FUNCTION_BLOCK Basic1_1 (* Basic Function Block Type *)
  (* Standard: 61499-2 *)
  (* Version 0.0, 1/4/2020, prana, nxtControl GmbH, Template *)
  PACKAGE Main;
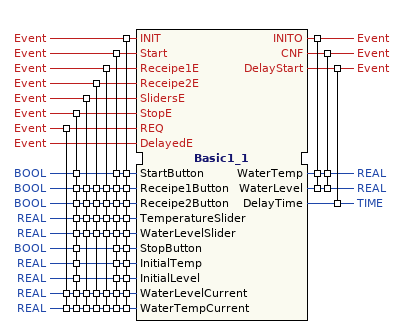
  EVENT_INPUT
    INIT WITH StartButton, Receipe1Button, Receipe2Button, TemperatureSlider, WaterLevelSlider, StopButton, InitialTemp, InitialLevel, WaterLevelCurrent, WaterTempCurrent;
    Start WITH StartButton, Receipe1Button, Receipe2Button, TemperatureSlider, WaterLevelSlider, StopButton, InitialTemp, InitialLevel, WaterLevelCurrent, WaterTempCurrent;
    Receipe1E WITH Receipe1Button, Receipe2Button, TemperatureSlider, WaterLevelSlider, WaterLevelCurrent, WaterTempCurrent; (* Initialization Request *)
    Receipe2E WITH Receipe1Button, Receipe2Button, TemperatureSlider, WaterLevelSlider, WaterLevelCurrent, WaterTempCurrent; (* Normal Execution Request *)
    SlidersE WITH Receipe1Button, Receipe2Button, TemperatureSlider, WaterLevelSlider, WaterLevelCurrent, WaterTempCurrent;
    StopE WITH StartButton, Receipe1Button, Receipe2Button, TemperatureSlider, WaterLevelSlider, StopButton, InitialTemp, InitialLevel, WaterLevelCurrent, WaterTempCurrent;
    REQ WITH WaterLevelCurrent, WaterTempCurrent;
    DelayedE;
  END_EVENT
  EVENT_OUTPUT
    INITO WITH WaterLevel, WaterTemp; (* Initialization Confirm *)
    CNF WITH WaterLevel, WaterTemp; (* Execution Confirmation *)
    DelayStart WITH DelayTime;
  END_EVENT
  VAR_INPUT
    StartButton : BOOL;
    Receipe1Button : BOOL; (* Input event qualifier *)
    Receipe2Button : BOOL;
    TemperatureSlider : REAL;
    WaterLevelSlider : REAL;
    StopButton : BOOL;
    InitialTemp : REAL;
    InitialLevel : REAL;
    WaterLevelCurrent : REAL;
    WaterTempCurrent : REAL;
  END_VAR
  VAR_OUTPUT
    WaterTemp : REAL;
    WaterLevel : REAL; (* Output event qualifier *)
    DelayTime : TIME;
  END_VAR
  VAR
    X1 : REAL := 160.50;
    Y1 : REAL := 50.00;
    X2 : REAL := 250.50;
    Y2 : REAL := 68.96;
    X3 : REAL := 351.50;
    Y3 : REAL := 64.32;
    X4 : REAL := 180.00;
    Y4 : REAL := 42.60;
    T1 : TIME := T#3s;
    T2 : TIME := T#2s;
  END_VAR
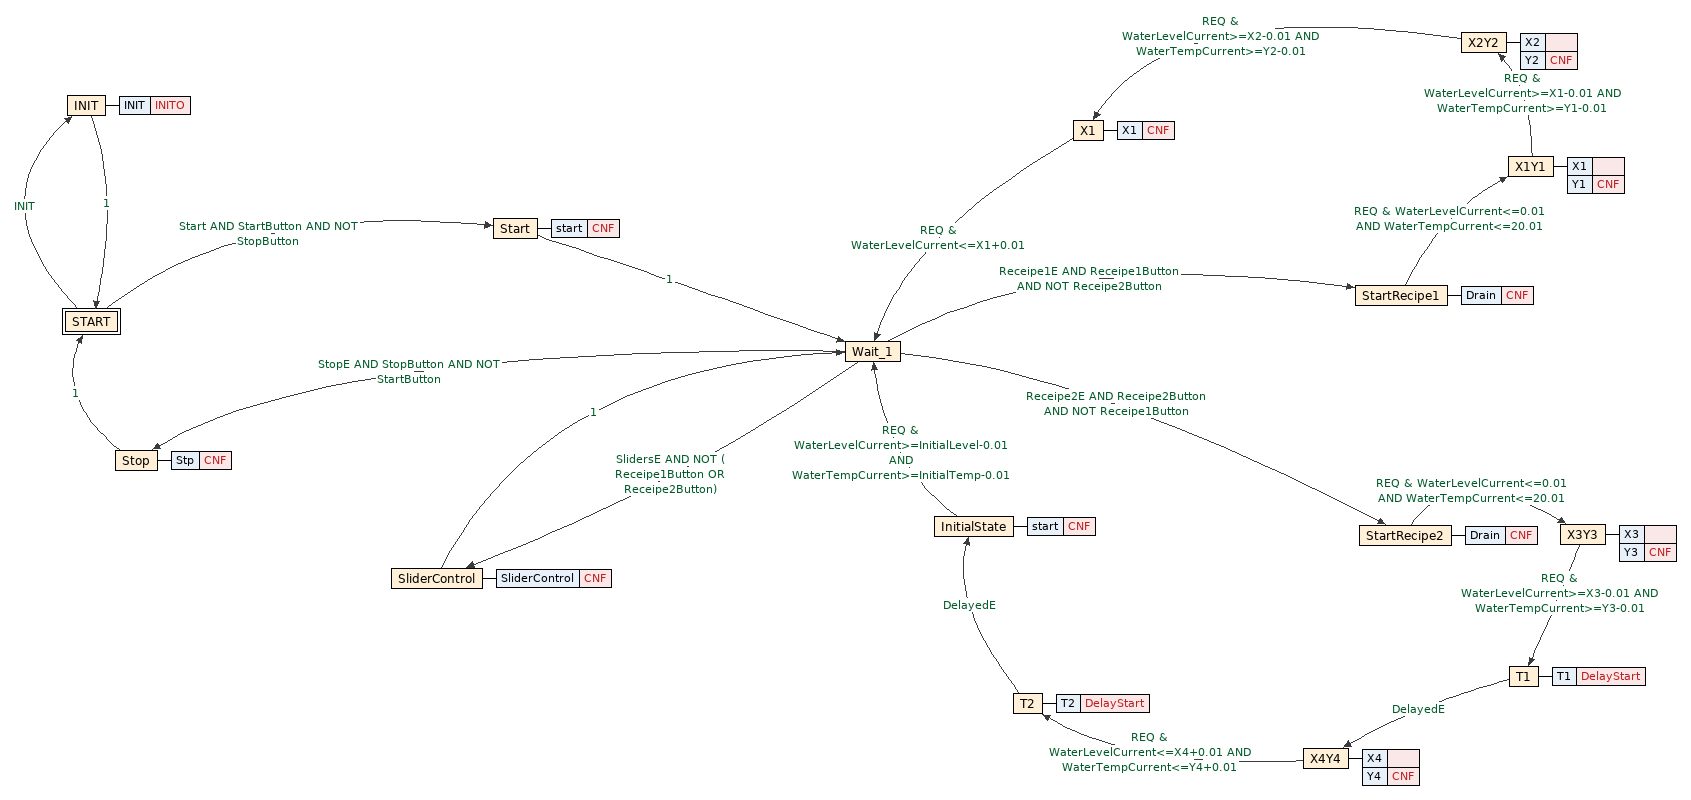
  EC_STATES
    START; (* Initial State *)
    SliderControl : SliderControl -> CNF;
    Start : start -> CNF;
    Wait_1;
    Stop : Stp -> CNF;
    INIT : INIT -> INITO;
    StartRecipe1 : Drain -> CNF;
    StartRecipe2 : Drain -> CNF;
    X1Y1 : X1, Y1 -> CNF;
    X2Y2 : X2, Y2 -> CNF;
    X1 : X1 -> CNF;
    X3Y3 : X3, Y3 -> CNF;
    T1 : T1 -> DelayStart;
    X4Y4 : X4, Y4 -> CNF;
    T2 : T2 -> DelayStart;
    InitialState : start -> CNF;
  END_STATES
  EC_TRANSITIONS
    Wait_1 TO SliderControl := SlidersE AND NOT ( Receipe1Button OR Receipe2Button);
    SliderControl TO Wait_1 := 1;
    START TO Start := Start AND StartButton AND NOT StopButton;
    Wait_1 TO Stop := StopE AND StopButton AND NOT StartButton;
    Stop TO START := 1;
    START TO INIT := INIT;
    INIT TO START := 1;
    StartRecipe1 TO X1Y1 := REQ & WaterLevelCurrent<=0.01 AND WaterTempCurrent<=20.01;
    X1Y1 TO X2Y2 := REQ & WaterLevelCurrent>=X1-0.01 AND WaterTempCurrent>=Y1-0.01;
    X3Y3 TO T1 := REQ & WaterLevelCurrent>=X3-0.01 AND WaterTempCurrent>=Y3-0.01;
    T1 TO X4Y4 := DelayedE;
    T2 TO InitialState := DelayedE;
    InitialState TO Wait_1 := REQ & WaterLevelCurrent>=InitialLevel-0.01 AND WaterTempCurrent>=InitialTemp-0.01;
    X2Y2 TO X1 := REQ & WaterLevelCurrent>=X2-0.01 AND WaterTempCurrent>=Y2-0.01;
    X1 TO Wait_1 := REQ & WaterLevelCurrent<=X1+0.01;
    Start TO Wait_1 := 1;
    Wait_1 TO StartRecipe1 := Receipe1E AND Receipe1Button AND NOT Receipe2Button;
    Wait_1 TO StartRecipe2 := Receipe2E AND Receipe2Button AND NOT Receipe1Button;
    StartRecipe2 TO X3Y3 := REQ & WaterLevelCurrent<=0.01 AND WaterTempCurrent<=20.01;
    X4Y4 TO T2 := REQ & WaterLevelCurrent<=X4+0.01 AND WaterTempCurrent<=Y4+0.01;
  END_TRANSITIONS
  ALGORITHM INIT IN ST: (* Initialization algorithm *)
;
  END_ALGORITHM
  ALGORITHM SliderControl IN ST:
WaterLevel := WaterLevelSlider;
WaterTemp := TemperatureSlider;
  END_ALGORITHM
  ALGORITHM start IN ST:
WaterLevel := InitialLevel;
WaterTemp := InitialTemp;
  END_ALGORITHM
  ALGORITHM Stp IN ST:
WaterLevel := 0;
WaterTemp := 0;
  END_ALGORITHM
  ALGORITHM Drain IN ST:
WaterLevel:=0;
WaterTemp:=0;
  END_ALGORITHM
  ALGORITHM X1 IN ST:
WaterLevel:=X1;
  END_ALGORITHM
  ALGORITHM Y1 IN ST:
WaterTemp:=Y1;
  END_ALGORITHM
  ALGORITHM X2 IN ST:
WaterLevel:=X2;
  END_ALGORITHM
  ALGORITHM Y2 IN ST:
WaterTemp:=Y2;
  END_ALGORITHM
  ALGORITHM X3 IN ST:
WaterLevel:=X3;
  END_ALGORITHM
  ALGORITHM X4 IN ST:
WaterLevel:=X4;
  END_ALGORITHM
  ALGORITHM Y3 IN ST:
WaterTemp:=Y3;
  END_ALGORITHM
  ALGORITHM Y4 IN ST:
WaterTemp:=Y4;
  END_ALGORITHM
  ALGORITHM T1 IN ST:
DelayTime:=T1;
  END_ALGORITHM
  ALGORITHM T2 IN ST:
DelayTime:=T2;
  END_ALGORITHM
END_FUNCTION_BLOCK
